Fanuc KAREL source: kb00040.KL

-- PROVISIONAL review KL for V1013-1; original PC SHA256 5a4949706cd3aa0a39288463fd84f5833338b98b006ebb3850a4d5ba41c6b5b4
-- Incomplete behavior may be omitted. Consult companion uncertainty JSON. Do not deploy.
PROGRAM KB00040
%NOLOCKGROUP
BEGIN
  -- UNRESOLVED_PC offsets 5-14; opcodes 3F,75
  -- UNRESOLVED_PC offsets 19-26; opcodes 9D,23
  -- UNRESOLVED_PC offsets 31-49; opcodes 27,22,2A,22,31
  -- UNRESOLVED_PC offsets 54-58; opcodes 7F
END KB00040
